(* IEC 61131-3 sources: Piper/PiperModuleTemplate, 3 files *)

(* ---- Cyclic.st ---- *)
(********************************************************************
 * COPYRIGHT --
 ********************************************************************
 * Program: PiperModuleTemplate
 * File: PiperModuleTemplateCyclic.st
 * Author: Josh
 * Created: October 03, 2013
 ********************************************************************
 * Implementation of program PiperModuleTemplate
 ********************************************************************)

PROGRAM _CYCLIC

	// Call PiperModuleInterface to interface with the rest of the machine
	PiperModuleInterface;

	//Put your code here

END_PROGRAM

(* ---- PiperInterface.st ---- *)
(********************************************************************
 * COPYRIGHT --
 ********************************************************************
 * Program: MachineProg
 * File: PiperModuleInterface.st
 * Author: Josh
 * Created: October 03, 2013
 ********************************************************************
 * Implementation of program MachineProg
 ********************************************************************)

ACTION PiperModuleInterface:

	//Give this module a name so it is easier to debug
	ModuleInterface.ModuleName:=	'Name';

	//Add a module to the Piper
	Module.ModuleInterface:=	ADR(ModuleInterface);
	Module.Piper:= 	ADR(gMachine);
	Module();

	// Handle any machine states that this module needs to respond to
	CASE ModuleInterface.PiperState OF
//		MACH_ST_BOOTING:
//		MACH_ST_CLEARING:
//		MACH_ST_STOPPED:
//		MACH_ST_STARTING:
//		MACH_ST_IDLE:
//		MACH_ST_SUSPENDED:
//		MACH_ST_EXECUTE:
//		MACH_ST_STOPPING:
//		MACH_ST_ABORTING:
//		MACH_ST_ABORTED:
//		MACH_ST_HOLDING:
//		MACH_ST_HELD:
//		MACH_ST_UNHOLDING:
//		MACH_ST_SUSPENDING:
//		MACH_ST_UNSUSPENDING:
//		MACH_ST_RESETTING:
//		MACH_ST_COMPLETING:
//		MACH_ST_COMPLETE:

		MACH_ST_BYPASSED:

		ELSE
			ModuleInterface.ModuleResponse:=	ModuleInterface.PiperState;

	END_CASE

END_ACTION

(* ---- PiperModule.var ---- *)
(********************************************************************
 * COPYRIGHT --
 ********************************************************************
 * Program: PiperModuleTemplate
 * File: PiperModuleTemplate.var
 * Author: Josh
 * Created: October 03, 2013
 ********************************************************************
 * Local variables of program PiperModuleTemplate
 ********************************************************************)
VAR
	ModuleInterface : Module_Interface_typ;
	Module : Piper_Module_Fub;
END_VAR
